(* IEC 61131-3 sources: Versio-VersionControlSystem/fixtures/projects/RefrigeratorControl_FBS/RefrigeratorControl.fbsproj/Device.device.xml.v3^/Plc Logic.plclogic.xml.v3^/Application.application.xml.v3^/Library/Alarm/GVLs, 1 file *)

(* ---- GVL_Alarm.gvl ---- *)
(* METADATA
{
	"v3Meta": {
		"objectGuid": "4686c4cd-f467-4000-9d56-feab29dfab29"
	}
}
*)
{attribute 'qualified_only'}
NAMESPACE GVL_Alarm
VAR_GLOBAL
	AlarmConstant : DINT := 3;
END_VAR
END_NAMESPACE
